// TIA Portal V19 export
// export: Created 2026-10-15T10:10:35.4045672Z, ExportSetting WithDefaults, DisplayName Totally Integrated Automation Portal, DisplayVersion V19, DisplayName TIA Portal Openness, DisplayVersion V19, DisplayName TIA Portal Version Control Interface, DisplayVersion V19, DisplayName STEP 7 Professional, DisplayVersion V19, DisplayName STEP 7 Safety, DisplayVersion V19, DisplayName WinCC Basic/Comfort/Advanced, DisplayVersion V19, DisplayName WinCC Unified, DisplayVersion V19
FUNCTION "ROLL_PB4" : Void   // FC16, SCL
{ S7_Optimized_Access := 'TRUE' }
VERSION : 0.1
// stored: AutoNumber true, IsIECCheckEnabled false, SetENOAutomatically false, UDAEnableTagReadback false
   VAR_TEMP
      r : Bool;
      a1 : Word;
      a2 : Word;
      activeDataBlock : Int;
      comparisonResults : Array[0..24] of Bool;
   END_VAR
BEGIN

   #r := FALSE;
   #a1 := W#16#0000;
   #a2 := W#16#0000;
   #activeDataBlock := 0;
   // PB4, STEP 5 network 1
   #a2 := #a1;
   #a1 := "ROLL_GetM"(FirstByte := 239, Width := 8);
   #a2 := #a1;
   #a1 := W#16#001E;
   #comparisonResults[0] := (WORD_TO_INT(#a2) = WORD_TO_INT(#a1));
   #r := #comparisonResults[0];
   "ROLL_State".M[23, 5] := #r;
   // PB4, STEP 5 network 2
   #a2 := #a1;
   #a1 := "ROLL_GetM"(FirstByte := 239, Width := 8);
   #a2 := #a1;
   #a1 := W#16#001F;
   #comparisonResults[1] := (WORD_TO_INT(#a2) = WORD_TO_INT(#a1));
   #r := #comparisonResults[1];
   "ROLL_State".M[23, 6] := #r;
   // PB4, STEP 5 network 3
   #a2 := #a1;
   #a1 := "ROLL_GetM"(FirstByte := 239, Width := 8);
   #a2 := #a1;
   #a1 := W#16#0023;
   #comparisonResults[2] := (WORD_TO_INT(#a2) = WORD_TO_INT(#a1));
   #r := #comparisonResults[2];
   "ROLL_State".M[24, 0] := #r;
   // PB4, STEP 5 network 4
   #a2 := #a1;
   #a1 := "ROLL_GetM"(FirstByte := 239, Width := 8);
   #a2 := #a1;
   #a1 := W#16#0024;
   #comparisonResults[3] := (WORD_TO_INT(#a2) = WORD_TO_INT(#a1));
   #r := #comparisonResults[3];
   "ROLL_State".M[24, 1] := #r;
   // PB4, STEP 5 network 5
   #a2 := #a1;
   #a1 := "ROLL_GetM"(FirstByte := 239, Width := 8);
   #a2 := #a1;
   #a1 := W#16#0025;
   #comparisonResults[4] := (WORD_TO_INT(#a2) = WORD_TO_INT(#a1));
   #r := #comparisonResults[4];
   "ROLL_State".M[24, 2] := #r;
   // PB4, STEP 5 network 6
   #a2 := #a1;
   #a1 := "ROLL_GetM"(FirstByte := 239, Width := 8);
   #a2 := #a1;
   #a1 := W#16#0026;
   #comparisonResults[5] := (WORD_TO_INT(#a2) = WORD_TO_INT(#a1));
   #r := #comparisonResults[5];
   "ROLL_State".M[24, 3] := #r;
   // PB4, STEP 5 network 7
   #a2 := #a1;
   #a1 := "ROLL_GetM"(FirstByte := 239, Width := 8);
   #a2 := #a1;
   #a1 := W#16#0027;
   #comparisonResults[6] := (WORD_TO_INT(#a2) = WORD_TO_INT(#a1));
   #r := #comparisonResults[6];
   "ROLL_State".M[24, 4] := #r;
   // PB4, STEP 5 network 8
   #a2 := #a1;
   #a1 := "ROLL_GetM"(FirstByte := 239, Width := 8);
   #a2 := #a1;
   #a1 := W#16#0032;
   #comparisonResults[7] := (WORD_TO_INT(#a2) = WORD_TO_INT(#a1));
   #r := #comparisonResults[7];
   "ROLL_State".M[25, 0] := #r;
   // PB4, STEP 5 network 9
   #a2 := #a1;
   #a1 := "ROLL_GetM"(FirstByte := 239, Width := 8);
   #a2 := #a1;
   #a1 := W#16#0033;
   #comparisonResults[8] := (WORD_TO_INT(#a2) = WORD_TO_INT(#a1));
   #r := #comparisonResults[8];
   "ROLL_State".M[25, 1] := #r;
   // PB4, STEP 5 network 10
   #a2 := #a1;
   #a1 := "ROLL_GetM"(FirstByte := 239, Width := 8);
   #a2 := #a1;
   #a1 := W#16#0034;
   #comparisonResults[9] := (WORD_TO_INT(#a2) = WORD_TO_INT(#a1));
   #r := #comparisonResults[9];
   "ROLL_State".M[25, 2] := #r;
   // PB4, STEP 5 network 11
   #a2 := #a1;
   #a1 := "ROLL_GetM"(FirstByte := 239, Width := 8);
   #a2 := #a1;
   #a1 := W#16#0035;
   #comparisonResults[10] := (WORD_TO_INT(#a2) = WORD_TO_INT(#a1));
   #r := #comparisonResults[10];
   "ROLL_State".M[25, 3] := #r;
   // PB4, STEP 5 network 12
   #a2 := #a1;
   #a1 := "ROLL_GetM"(FirstByte := 239, Width := 8);
   #a2 := #a1;
   #a1 := W#16#0037;
   #comparisonResults[11] := (WORD_TO_INT(#a2) = WORD_TO_INT(#a1));
   #r := #comparisonResults[11];
   "ROLL_State".M[25, 4] := #r;
   // PB4, STEP 5 network 13
   #a2 := #a1;
   #a1 := "ROLL_GetM"(FirstByte := 239, Width := 8);
   #a2 := #a1;
   #a1 := W#16#0038;
   #comparisonResults[12] := (WORD_TO_INT(#a2) = WORD_TO_INT(#a1));
   #r := #comparisonResults[12];
   "ROLL_State".M[25, 5] := #r;
   // PB4, STEP 5 network 14
   #a2 := #a1;
   #a1 := "ROLL_GetM"(FirstByte := 239, Width := 8);
   #a2 := #a1;
   #a1 := W#16#0039;
   #comparisonResults[13] := (WORD_TO_INT(#a2) = WORD_TO_INT(#a1));
   #r := #comparisonResults[13];
   "ROLL_State".M[25, 6] := #r;
   // PB4, STEP 5 network 15
   #a2 := #a1;
   #a1 := "ROLL_GetM"(FirstByte := 239, Width := 8);
   #a2 := #a1;
   #a1 := W#16#003A;
   #comparisonResults[14] := (WORD_TO_INT(#a2) = WORD_TO_INT(#a1));
   #r := #comparisonResults[14];
   "ROLL_State".M[25, 7] := #r;
   // PB4, STEP 5 network 16
   #a2 := #a1;
   #a1 := "ROLL_GetM"(FirstByte := 239, Width := 8);
   #a2 := #a1;
   #a1 := W#16#003C;
   #comparisonResults[15] := (WORD_TO_INT(#a2) = WORD_TO_INT(#a1));
   #r := #comparisonResults[15];
   "ROLL_State".M[26, 0] := #r;
   // PB4, STEP 5 network 17
   #a2 := #a1;
   #a1 := "ROLL_GetM"(FirstByte := 239, Width := 8);
   #a2 := #a1;
   #a1 := W#16#003D;
   #comparisonResults[16] := (WORD_TO_INT(#a2) = WORD_TO_INT(#a1));
   #r := #comparisonResults[16];
   "ROLL_State".M[26, 1] := #r;
   // PB4, STEP 5 network 18
   #a2 := #a1;
   #a1 := "ROLL_GetM"(FirstByte := 239, Width := 8);
   #a2 := #a1;
   #a1 := W#16#003E;
   #comparisonResults[17] := (WORD_TO_INT(#a2) = WORD_TO_INT(#a1));
   #r := #comparisonResults[17];
   "ROLL_State".M[26, 2] := #r;
   // PB4, STEP 5 network 19
   #a2 := #a1;
   #a1 := "ROLL_GetM"(FirstByte := 239, Width := 8);
   #a2 := #a1;
   #a1 := W#16#003F;
   #comparisonResults[18] := (WORD_TO_INT(#a2) = WORD_TO_INT(#a1));
   #r := #comparisonResults[18];
   "ROLL_State".M[26, 3] := #r;
   // PB4, STEP 5 network 20
   #a2 := #a1;
   #a1 := "ROLL_GetM"(FirstByte := 239, Width := 8);
   #a2 := #a1;
   #a1 := W#16#0041;
   #comparisonResults[19] := (WORD_TO_INT(#a2) = WORD_TO_INT(#a1));
   #r := #comparisonResults[19];
   "ROLL_State".M[26, 5] := #r;
   // PB4, STEP 5 network 21
   #a2 := #a1;
   #a1 := "ROLL_GetM"(FirstByte := 239, Width := 8);
   #a2 := #a1;
   #a1 := W#16#0042;
   #comparisonResults[20] := (WORD_TO_INT(#a2) = WORD_TO_INT(#a1));
   #r := #comparisonResults[20];
   "ROLL_State".M[26, 6] := #r;
   // PB4, STEP 5 network 22
   #a2 := #a1;
   #a1 := "ROLL_GetM"(FirstByte := 239, Width := 8);
   #a2 := #a1;
   #a1 := W#16#0045;
   #comparisonResults[21] := (WORD_TO_INT(#a2) = WORD_TO_INT(#a1));
   #r := #comparisonResults[21];
   "ROLL_State".M[27, 1] := #r;
   // PB4, STEP 5 network 23
   #a2 := #a1;
   #a1 := "ROLL_GetM"(FirstByte := 239, Width := 8);
   #a2 := #a1;
   #a1 := W#16#0048;
   #comparisonResults[22] := (WORD_TO_INT(#a2) = WORD_TO_INT(#a1));
   #r := #comparisonResults[22];
   "ROLL_State".M[27, 4] := #r;
   // PB4, STEP 5 network 24
   #a2 := #a1;
   #a1 := "ROLL_GetM"(FirstByte := 239, Width := 8);
   #a2 := #a1;
   #a1 := W#16#0049;
   #comparisonResults[23] := (WORD_TO_INT(#a2) = WORD_TO_INT(#a1));
   #r := #comparisonResults[23];
   "ROLL_State".M[27, 5] := #r;
   // PB4, STEP 5 network 25
   #a2 := #a1;
   #a1 := "ROLL_GetM"(FirstByte := 239, Width := 8);
   #a2 := #a1;
   #a1 := W#16#0063;
   #comparisonResults[24] := (WORD_TO_INT(#a2) = WORD_TO_INT(#a1));
   #r := #comparisonResults[24];
   "ROLL_State".M[27, 7] := #r;
   // PB4, STEP 5 network 26
   RETURN;
END_FUNCTION
